# EPICS substitutions: evrIoc/Db/patternSimXL04.substitutions
# ESIM Pattern records (from EVG) to EVR:
file evrPatternTestBsa.db {
  pattern { EIOC  ,  DEVICE }
	  { IOC:XX04:1  ,ESIM:XX04:1  }
}

# EVG EDEF checking simulation for Modifier5/ bsa enable/disable:
file bsaProcTestAll_event.db {
  pattern {  DEVICE,     LOC     }
	      { ESIM:XX04:1, SYS0    }
}
